// TIA Portal V19 export
FUNCTION_BLOCK "AUTO_HEATING_SELECTION"   // FB13, LAD
{ S7_Optimized_Access := 'TRUE' }
// COOLING TO HEAT
// stored: MemoryReserve 100, SetENOAutomatically false
   VAR_INPUT
      AUTO : Bool;
      RUNNING : Bool;
      CONTROL_MODE : Int;
      TEMP_PV : Real;
      HEAT_RUNNING : Bool;
      HEAT_UCH_MIN_SP : Real;
      HEAT_UCH_MAX_SP : Real;
      HEAT_CH_MIN_SP : Real;
      HEAT_CH_MAX_SP : Real;
      HEAT_CT_MIN_SP : Real;
      HEAT_CT_MAX_SP : Real;
      HEAT_HW_MIN_SP : Real;
      HEAT_HW_MAX_SP : Real;
   END_VAR
   VAR_OUTPUT
      UCHWS_CMD : Bool;
      CHWS_CMD : Bool;
      CTS_CMD : Bool;
      HWS_CMD : Bool;
      UTILITY_SEL : Int;
   END_VAR
   VAR
      UCHWS { S7_SetPoint := 'True'} : Bool;
      CHWS : Bool;
      CTS : Bool;
      HWS : Bool;
   END_VAR
   VAR_TEMP   // added for the SCL form of the ladder/FBD networks
      _w1 : Bool;
   END_VAR
BEGIN

REGION Network 1: HEATING
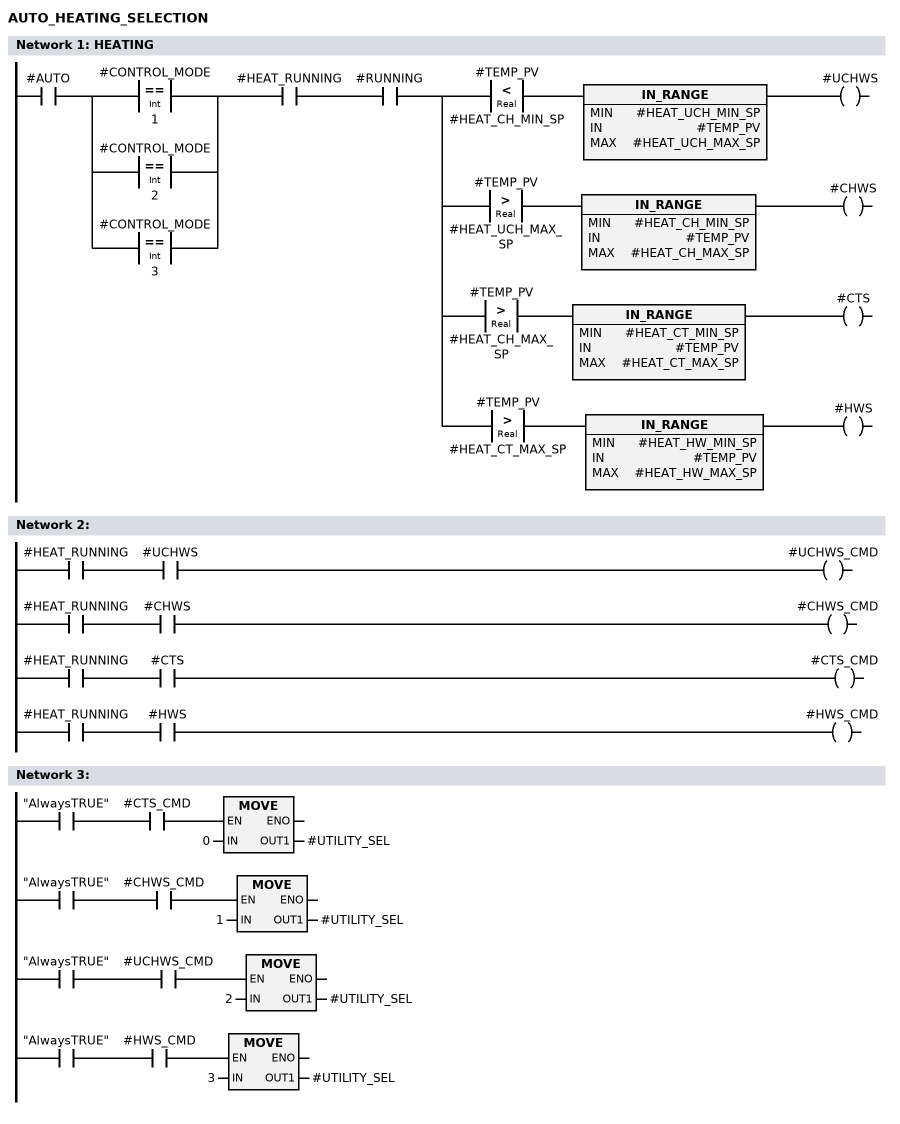
   RUNG wire#powerrail
      Contact( #AUTO )
      wire#w1
      { S7_Templates := "SrcType := Int" } EQ_Contact(in1 := #CONTROL_MODE, in2 := 1)
      wire#w2
      Contact( #HEAT_RUNNING )
      Contact( #RUNNING )
      wire#w3
      { S7_Templates := "SrcType := Real" } LT_Contact(in1 := #TEMP_PV, in2 := #HEAT_CH_MIN_SP)
      { S7_Templates := "SrcType := Real" } InRange(min := #HEAT_UCH_MIN_SP, in := #TEMP_PV, max := #HEAT_UCH_MAX_SP)
      Coil( #UCHWS )
   END_RUNG
   RUNG wire#w1
      { S7_Templates := "SrcType := Int" } EQ_Contact(in1 := #CONTROL_MODE, in2 := 2)
   END_RUNG wire#w2
   RUNG wire#w1
      { S7_Templates := "SrcType := Int" } EQ_Contact(in1 := #CONTROL_MODE, in2 := 3)
   END_RUNG wire#w2
   RUNG wire#w3
      { S7_Templates := "SrcType := Real" } GT_Contact(in1 := #TEMP_PV, in2 := #HEAT_UCH_MAX_SP)
      { S7_Templates := "SrcType := Real" } InRange(min := #HEAT_CH_MIN_SP, in := #TEMP_PV, max := #HEAT_CH_MAX_SP)
      Coil( #CHWS )
   END_RUNG
   RUNG wire#w3
      { S7_Templates := "SrcType := Real" } GT_Contact(in1 := #TEMP_PV, in2 := #HEAT_CH_MAX_SP)
      { S7_Templates := "SrcType := Real" } InRange(min := #HEAT_CT_MIN_SP, in := #TEMP_PV, max := #HEAT_CT_MAX_SP)
      Coil( #CTS )
   END_RUNG
   RUNG wire#w3
      { S7_Templates := "SrcType := Real" } GT_Contact(in1 := #TEMP_PV, in2 := #HEAT_CT_MAX_SP)
      { S7_Templates := "SrcType := Real" } InRange(min := #HEAT_HW_MIN_SP, in := #TEMP_PV, max := #HEAT_HW_MAX_SP)
      Coil( #HWS )
   END_RUNG
   // the same network as SCL:
   #_w1 := #AUTO AND ((#CONTROL_MODE = 1) OR (#CONTROL_MODE = 2) OR (#CONTROL_MODE = 3)) AND #HEAT_RUNNING AND #RUNNING;
   #UCHWS := #_w1 AND (#TEMP_PV < #HEAT_CH_MIN_SP) AND (#HEAT_UCH_MIN_SP <= #TEMP_PV) AND (#TEMP_PV <= #HEAT_UCH_MAX_SP);
   #CHWS := #_w1 AND (#TEMP_PV > #HEAT_UCH_MAX_SP) AND (#HEAT_CH_MIN_SP <= #TEMP_PV) AND (#TEMP_PV <= #HEAT_CH_MAX_SP);
   #CTS := #_w1 AND (#TEMP_PV > #HEAT_CH_MAX_SP) AND (#HEAT_CT_MIN_SP <= #TEMP_PV) AND (#TEMP_PV <= #HEAT_CT_MAX_SP);
   #HWS := #_w1 AND (#TEMP_PV > #HEAT_CT_MAX_SP) AND (#HEAT_HW_MIN_SP <= #TEMP_PV) AND (#TEMP_PV <= #HEAT_HW_MAX_SP);
END_REGION

REGION Network 2
   RUNG wire#powerrail
      Contact( #HEAT_RUNNING )
      Contact( #UCHWS )
      Coil( #UCHWS_CMD )
   END_RUNG
   RUNG wire#powerrail
      Contact( #HEAT_RUNNING )
      Contact( #CHWS )
      Coil( #CHWS_CMD )
   END_RUNG
   RUNG wire#powerrail
      Contact( #HEAT_RUNNING )
      Contact( #CTS )
      Coil( #CTS_CMD )
   END_RUNG
   RUNG wire#powerrail
      Contact( #HEAT_RUNNING )
      Contact( #HWS )
      Coil( #HWS_CMD )
   END_RUNG
   // the same network as SCL:
   #UCHWS_CMD := #HEAT_RUNNING AND #UCHWS;
   #CHWS_CMD := #HEAT_RUNNING AND #CHWS;
   #CTS_CMD := #HEAT_RUNNING AND #CTS;
   #HWS_CMD := #HEAT_RUNNING AND #HWS;
END_REGION

REGION Network 3
   RUNG wire#powerrail
      Contact( "AlwaysTRUE" )
      Contact( #CTS_CMD )
      Move(in := 0, out1 => #UTILITY_SEL)
   END_RUNG
   RUNG wire#powerrail
      Contact( "AlwaysTRUE" )
      Contact( #CHWS_CMD )
      Move(in := 1, out1 => #UTILITY_SEL)
   END_RUNG
   RUNG wire#powerrail
      Contact( "AlwaysTRUE" )
      Contact( #UCHWS_CMD )
      Move(in := 2, out1 => #UTILITY_SEL)
   END_RUNG
   RUNG wire#powerrail
      Contact( "AlwaysTRUE" )
      Contact( #HWS_CMD )
      Move(in := 3, out1 => #UTILITY_SEL)
   END_RUNG
   // the same network as SCL:
   IF "AlwaysTRUE" AND #CTS_CMD THEN #UTILITY_SEL := 0; END_IF;
   IF "AlwaysTRUE" AND #CHWS_CMD THEN #UTILITY_SEL := 1; END_IF;
   IF "AlwaysTRUE" AND #UCHWS_CMD THEN #UTILITY_SEL := 2; END_IF;
   IF "AlwaysTRUE" AND #HWS_CMD THEN #UTILITY_SEL := 3; END_IF;
END_REGION
END_FUNCTION_BLOCK
